PROGRAM MAIN
VAR
	fbKessel : FB_Kessel;
END_VAR

// Ein Aufruf pro Task-Zyklus (Zykluszeit z. B. 100 ms).
fbKessel();

END_PROGRAM

(* stored: Version 1.1.0.1, ProductVersion 3.1.4024.32
   POU MAIN: Id {3B2C8D4E-5F60-4B7C-9D8E-0F1A2B3C4D5E}, SpecialFunc None *)
